// TIA Portal V21 export
TYPE "UDT_Motor"
TITLE = Motor data
   STRUCT
      Enable : Bool;   // Release from the line control
      Running : Bool;   // Feedback: motor is running
      Fault : Bool;   // Motor protection tripped
      SpeedSetpoint : Real := 1450.0;   // Speed setpoint in rpm
      ActualSpeed : Real;   // Measured speed in rpm
      RunTime : Time := T#0MS;   // Accumulated run time
      StartCount : DInt := 0;   // Number of starts
   END_STRUCT;
END_TYPE
